// TIA Portal V19 export
// export: Created 2026-10-15T09:44:23.2692016Z, ExportSetting WithDefaults, DisplayName Totally Integrated Automation Portal, DisplayVersion V19, DisplayName TIA Portal Openness, DisplayVersion V19, DisplayName TIA Portal Version Control Interface, DisplayVersion V19, DisplayName STEP 7 Professional, DisplayVersion V19, DisplayName STEP 7 Safety, DisplayVersion V19, DisplayName WinCC Basic/Comfort/Advanced, DisplayVersion V19, DisplayName WinCC Unified, DisplayVersion V19
FUNCTION "ROLL_FB90" : Void   // FC12, SCL
{ S7_Optimized_Access := 'TRUE' }
VERSION : 0.1
// stored: AutoNumber true, IsIECCheckEnabled false, SetENOAutomatically false, UDAEnableTagReadback false
BEGIN

   "ROLL_State".M[110, 0] := ("ROLL_DB205".DW[5] AND W#16#0FFF) <> W#16#0000;
   "ROLL_State".M[110, 1] := ("ROLL_DB205".DW[17] AND W#16#0FFF) <> W#16#0000;
   "ROLL_State".M[110, 2] := ("ROLL_DB205".DW[25] AND W#16#0FFF) <> W#16#0000;
   "ROLL_State".M[110, 3] := ("ROLL_DB205".DW[33] AND W#16#0FFF) <> W#16#0000;
   "ROLL_State".M[111, 0] := "ROLL_DB205".DW[37] = W#16#0001;
   "ROLL_State".M[111, 1] := "ROLL_DB205".DW[37] = W#16#0002;
   "ROLL_State".M[111, 2] := "ROLL_DB205".DW[37] = W#16#0003;
   "ROLL_State".M[111, 5] := "ROLL_DB205".DW[37] = W#16#0004;
   "ROLL_State".M[111, 3] := "ROLL_DB205".DW[41] = W#16#0001;
   "ROLL_State".M[111, 4] := "ROLL_DB205".DW[13] = W#16#0001;
   "ROLL_SetMWord"(FirstByte := 250,
                   Value := W#16#0000);
END_FUNCTION
